(* IEC 61131-3 sources: NachHouse_TST/ExamplesCustomLogin/AutoLogin, 2 files *)

(* ---- AutoLogin.ST ---- *)
VAR_GLOBAL
  CustomizedLoginPage AT %S355.1 : BOOL := true;
END_VAR

VAR_GLOBAL RETAIN

END_VAR

VAR_GLOBAL

END_VAR

(* ---- prgMain.ST ---- *)
PROGRAM prgMain
  VAR
    a : UINT;
  END_VAR

  a := a + 1;

END_PROGRAM
